FUNCTION F_SealPass : BOOL
VAR_INPUT
    Image : ITcVnImage;
END_VAR
VAR_OUTPUT
    ResultCode : HRESULT;
    BrightSamples : UINT;
END_VAR
VAR
    Pixel : TcVnVector4_LREAL;
    SampleIndex : UDINT;
END_VAR

// Five sample points from the Cartesian centre line of the supplied 160 x 100 frames.
ResultCode := 0;
BrightSamples := 0;
FOR SampleIndex := 0 TO 4 DO
    ResultCode := F_VN_GetPixel(Image, Pixel, 80, 26 + 12 * SampleIndex, ResultCode);
    IF (ResultCode >= 0) AND (Pixel[0] >= 200) THEN
        BrightSamples := BrightSamples + 1;
    END_IF
END_FOR
F_SealPass := (ResultCode >= 0) AND (BrightSamples >= 4);

END_FUNCTION

(* stored: Version 1.1.0.1
   POU F_SealPass: Id {CFA70A26-15B3-4CD7-831F-930C68FCB5D2} *)
